FUNCTION_BLOCK FB_ConveyorStarter (* Migrated from IEC 61131-3 ST *)
  (* Standard: 61499-2 *)
  (* Version 1.0, 2026-11-06, st2fb *)
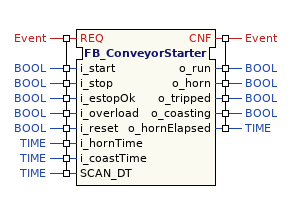
  EVENT_INPUT
    REQ WITH i_start, i_stop, i_estopOk, i_overload, i_reset, i_hornTime, i_coastTime, SCAN_DT;
  END_EVENT
  EVENT_OUTPUT
    CNF WITH o_run, o_horn, o_tripped, o_coasting, o_hornElapsed;
  END_EVENT
  VAR_INPUT
    i_start : BOOL;
    i_stop : BOOL;
    i_estopOk : BOOL;
    i_overload : BOOL;
    i_reset : BOOL;
    i_hornTime : TIME;
    i_coastTime : TIME;
    SCAN_DT : TIME;
  END_VAR
  VAR_OUTPUT
    o_run : BOOL;
    o_horn : BOOL;
    o_tripped : BOOL;
    o_coasting : BOOL;
    o_hornElapsed : TIME;
  END_VAR
  VAR
    statRunRequest : BOOL;
    statTrip : BOOL;
    statHornPreset : TIME;
    statCoastPreset : TIME;
    tempPermit : BOOL;
    ST2FB_NOW : TIME;
    statStartEdge_CLK : BOOL;
    statStartEdge_Q : BOOL;
    statStartEdge_M : BOOL;
    statHornTimer_IN : BOOL;
    statHornTimer_PT : TIME;
    statHornTimer_Q : BOOL;
    statHornTimer_ET : TIME;
    statHornTimer_STATE : INT;
    statHornTimer_PREV_IN : BOOL;
    statHornTimer_START_TIME : TIME;
    statCoastTimer_IN : BOOL;
    statCoastTimer_PT : TIME;
    statCoastTimer_Q : BOOL;
    statCoastTimer_ET : TIME;
    statCoastTimer_STATE : INT;
    statCoastTimer_PREV_IN : BOOL;
    statCoastTimer_START_TIME : TIME;
  END_VAR
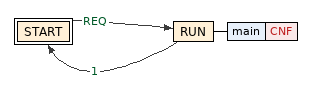
  EC_STATES
    START;
    RUN : main -> CNF;
  END_STATES
  EC_TRANSITIONS
    START TO RUN := REQ;
    RUN TO START := 1;
  END_TRANSITIONS
  ALGORITHM main IN ST:
ST2FB_NOW := ST2FB_NOW + SCAN_DT;
IF i_overload OR NOT i_estopOk THEN
  statTrip := TRUE;
ELSIF i_reset THEN
  statTrip := FALSE;
END_IF;
tempPermit := i_estopOk AND NOT statTrip;

IF NOT statRunRequest THEN
  statHornPreset := i_hornTime;
END_IF;
IF o_run THEN
  statCoastPreset := i_coastTime;
END_IF;
statStartEdge_CLK := i_start;
statStartEdge_Q := statStartEdge_CLK AND NOT statStartEdge_M;
statStartEdge_M := statStartEdge_CLK;
IF i_stop OR NOT tempPermit THEN
  statRunRequest := FALSE;
ELSIF statStartEdge_Q THEN
  statRunRequest := TRUE;
END_IF;

statHornTimer_IN := statRunRequest;
statHornTimer_PT := statHornPreset;
IF (statHornTimer_STATE = 0) AND NOT statHornTimer_PREV_IN AND statHornTimer_IN THEN
  statHornTimer_STATE := 1;
  statHornTimer_Q := FALSE;
  statHornTimer_START_TIME := ST2FB_NOW;
ELSE
  IF NOT statHornTimer_IN THEN
    statHornTimer_ET := T#0s;
    statHornTimer_Q := FALSE;
    statHornTimer_STATE := 0;
  ELSIF statHornTimer_STATE = 1 THEN
    IF statHornTimer_START_TIME + statHornTimer_PT <= ST2FB_NOW THEN
      statHornTimer_STATE := 2;
      statHornTimer_Q := TRUE;
      statHornTimer_ET := statHornTimer_PT;
    ELSE
      statHornTimer_ET := ST2FB_NOW - statHornTimer_START_TIME;
    END_IF;
  END_IF;
END_IF;
statHornTimer_PREV_IN := statHornTimer_IN;
o_hornElapsed := statHornTimer_ET;
o_horn := statRunRequest AND NOT statHornTimer_Q;
o_run := statRunRequest AND statHornTimer_Q;

statCoastTimer_IN := o_run;
statCoastTimer_PT := statCoastPreset;
IF (statCoastTimer_STATE = 0) AND statCoastTimer_PREV_IN AND NOT statCoastTimer_IN THEN
  statCoastTimer_STATE := 1;
  statCoastTimer_START_TIME := ST2FB_NOW;
ELSE
  IF statCoastTimer_IN THEN
    statCoastTimer_ET := T#0s;
    statCoastTimer_STATE := 0;
  ELSIF statCoastTimer_STATE = 1 THEN
    IF statCoastTimer_START_TIME + statCoastTimer_PT <= ST2FB_NOW THEN
      statCoastTimer_STATE := 2;
      statCoastTimer_ET := statCoastTimer_PT;
    ELSE
      statCoastTimer_ET := ST2FB_NOW - statCoastTimer_START_TIME;
    END_IF;
  END_IF;
END_IF;
statCoastTimer_Q := statCoastTimer_IN OR (statCoastTimer_STATE = 1);
statCoastTimer_PREV_IN := statCoastTimer_IN;
o_coasting := statCoastTimer_Q AND NOT o_run;
o_tripped := statTrip;
  END_ALGORITHM
END_FUNCTION_BLOCK
